Universal Robots URScript: T003_mistralai_Mistral-Large-3-675B-Instruct-2512-NVFP4_edit_perf_rep1.urscript

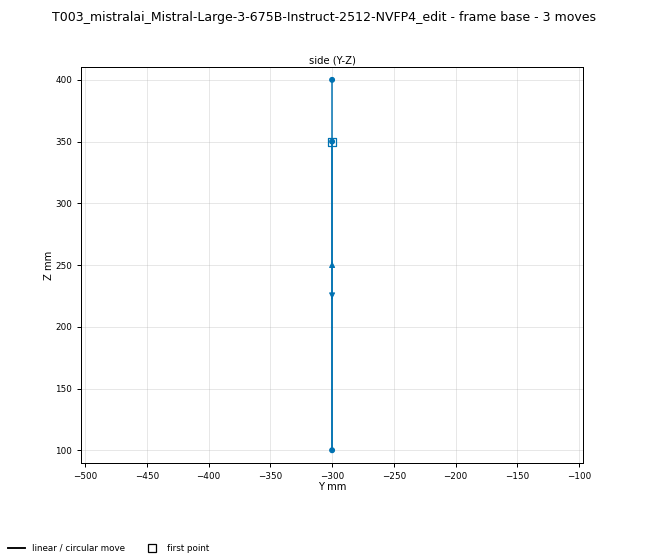
[picture p0: tool path of T003_mistralai_Mistral-Large-3-675B-Instruct-2512-NVFP4_edit_perf_rep1.urscript in frame base, 3 of 8 moves have a stored position in this frame; points joined in program order, loops and branches not executed]
def task_T003():
  # Safety check
  if (get_digital_in(0) == True):
    popup("E-Stop active — aborting program.", error=True)
    halt
  end

  # Home position - increased acceleration
  movej([0.0000, -1.5708, 1.5708, -1.5708, -1.5708, 0.0000], a=2.0000, v=1.0000)

  # Pre-calculate pallet positions
  pallet_origin = p[0.500000, 0.300000, 0.400000, 0.0000, 3.1416, 0.0000]
  positions = [
    pallet_origin,
    pallet_origin * p[0.0, 0.200, 0.0, 0.0, 0.0, 0.0],
    pallet_origin * p[0.200, 0.0, 0.0, 0.0, 0.0, 0.0],
    pallet_origin * p[0.200, 0.200, 0.0, 0.0, 0.0, 0.0]
  ]

  # Pick and place cycle for all 4 positions
  for i in range(4):
    # Approach conveyor pick - optimized path
    movel(p[0.500000, -0.300000, 0.350000, 0.0000, 3.1416, 0.0000], a=2.0000, v=0.3000, r=0.0200)

    # Descend to pick - faster descent
    movel(p[0.500000, -0.300000, 0.100000, 0.0000, 3.1416, 0.0000], a=1.0000, v=0.1500)

    # Gripper CLOSE - parallel with motion
    set_digital_out(0, True)
    sleep(0.1000)  # Reduced settle time

    # Lift from conveyor - increased speed
    movel(p[0.500000, -0.300000, 0.400000, 0.0000, 3.1416, 0.0000], a=1.5000, v=0.2500, r=0.0150)

    # Transit to pallet - max speed
    movel(positions[i], a=2.0000, v=0.3000, r=0.0200)

    # Descend to place - faster descent
    movel(positions[i] * p[0.0, 0.0, -0.280, 0.0, 0.0, 0.0], a=1.0000, v=0.1500)

    # Gripper OPEN - parallel with motion
    set_digital_out(0, False)
    sleep(0.1000)  # Reduced settle time

    # Retract above pallet - increased speed
    movel(positions[i], a=1.5000, v=0.2500, r=0.0100)

    # Return to home after last position
    if (i == 3):
      movej([0.0000, -1.5708, 1.5708, -1.5708, -1.5708, 0.0000], a=2.0000, v=1.0000)
    end
  end
end

task_T003()
